Fanuc KAREL source: kt00618.KL

PROGRAM KT00618
%NOLOCKGROUP
VAR
B1:BOOLEAN;B2:BOOLEAN;OUT:BOOLEAN
BEGIN
--
--
B1=TRUE
B2=FALSE
B1=TRUE
B2=FALSE
OUT=(NOT B1)
END KT00618
